// TIA Portal project "s15_motor" (V21)

(* hardware
DEVICE "S7-1500/ET200MP station_1"  S7-1500 station
   slot 0: "Rail_0"  Rack  6ES7 590-1***0-0AA0
   slot 1: "MOTORPLC"  CPU 1511-1 PN  6ES7 511-1AL03-0AB0  V4.1
      slot 3: "CPU display_1"  6ES7591-1AA00-0AA0
      slot 32768: "PROFINET interface_1"  X1
         slot 32769: "Port_1"  X1 P1
         slot 32770: "Port_2"  X1 P2
      slot 34817: "Virtual CP interface port_1"  Virtual CP interface port  Virtual CP interface port FW V4.1
*)

// ===== PLC "MOTORPLC"  CPU 1511-1 PN =====

VAR_GLOBAL   // PLC tag table "Default tag table"
   "StartPB" AT %I0.0 : Bool;   // start button, normally open
   "StopPB" AT %I0.1 : Bool;   // stop button, normally closed
   "Guard" AT %I0.2 : Bool;   // guard closed
   "MotorLadOut" AT %Q0.0 : Bool;
   "MotorSclOut" AT %Q0.1 : Bool;
END_VAR

DATA_BLOCK "MotorData"   // DB1
{ S7_Optimized_Access := 'TRUE' }
VERSION : 0.1
   VAR
      starts : Int;
      runTime : Time;
   END_VAR
BEGIN
END_DATA_BLOCK

DATA_BLOCK "MotorLAD_DB"   // DB2
{ S7_Optimized_Access := 'TRUE' }
VERSION : 0.1
// stored: InstanceOfName MotorLAD
"MotorLAD"
BEGIN
END_DATA_BLOCK

DATA_BLOCK "MotorSCL_DB"   // DB3
{ S7_Optimized_Access := 'TRUE' }
VERSION : 0.1
// stored: InstanceOfName MotorSCL
"MotorSCL"
BEGIN
END_DATA_BLOCK

FUNCTION_BLOCK "MotorLAD"   // FB1, LAD
{ S7_Optimized_Access := 'TRUE' }
VERSION : 0.1
   VAR_INPUT
      start : Bool;
      stop : Bool;
      interlock : Bool;
   END_VAR
   VAR_OUTPUT
      motor : Bool;
   END_VAR
   VAR
      run : Bool;
      runEdge : Bool;
      delay : TON_TIME;
   END_VAR
   VAR_TEMP   // added for the SCL form of the ladder/FBD networks
      _w1 : Bool;
   END_VAR
BEGIN

REGION Network 1
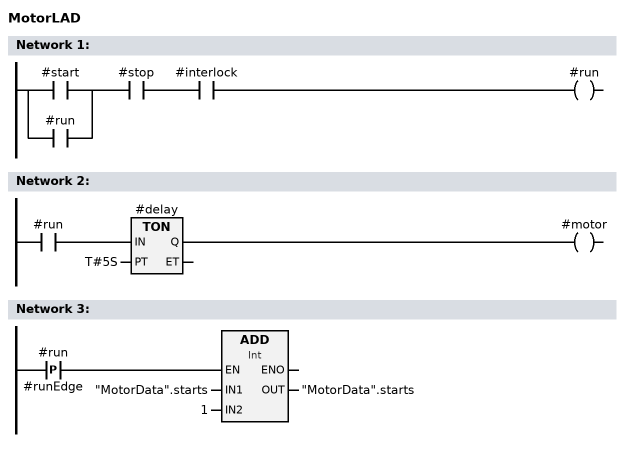
   RUNG wire#powerrail
      Contact( #start )
      wire#w1
      Contact( #stop )
      Contact( #interlock )
      Coil( #run )
   END_RUNG
   RUNG wire#powerrail
      Contact( #run )
   END_RUNG wire#w1
   // the same network as SCL:
   #run := (#start OR #run) AND #stop AND #interlock;
END_REGION

REGION Network 2
   #delay(IN := #run, PT := T#5S);   // TON
   #motor := #delay.Q;
END_REGION

REGION Network 3
   RUNG wire#powerrail
      P_Contact(operand := #run, bit := #runEdge)
      { S7_Templates := "SrcType := Int" } Add(in1 := "MotorData".starts, in2 := 1, out => "MotorData".starts)
   END_RUNG
   // the same network as SCL:
   #_w1 := #run AND NOT #runEdge;   // rising edge of #run
   #runEdge := #run;
   IF #_w1 THEN "MotorData".starts := "MotorData".starts + 1; END_IF;
END_REGION
END_FUNCTION_BLOCK

FUNCTION_BLOCK "MotorSCL"   // FB2, SCL
{ S7_Optimized_Access := 'TRUE' }
VERSION : 0.1
   VAR_INPUT
      start : Bool;
      stop : Bool;
      interlock : Bool;
   END_VAR
   VAR_OUTPUT
      motor : Bool;
   END_VAR
   VAR
      run : Bool;
      runOld : Bool;
      delay : TON_TIME;
   END_VAR
BEGIN
       // seal-in with interlock
       #run := (#start OR #run) AND #stop AND #interlock;
       // start delay
       #delay(IN := #run,
              PT := T#5S);
       #motor := #delay.Q;
       // count the starts
       IF #run AND NOT #runOld THEN
           "MotorData".starts := "MotorData".starts + 1;
       END_IF;
       #runOld := #run;
END_FUNCTION_BLOCK

ORGANIZATION_BLOCK "Main"   // OB1, LAD, ProgramCycle
TITLE = "Main Program Sweep (Cycle)"
{ S7_Optimized_Access := 'TRUE' }
VERSION : 0.1
   VAR_INPUT
      Initial_Call : Bool;   // Initial call of this OB
      Remanence : Bool;   // =True, if remanent data are available
   END_VAR
BEGIN

REGION Network 1
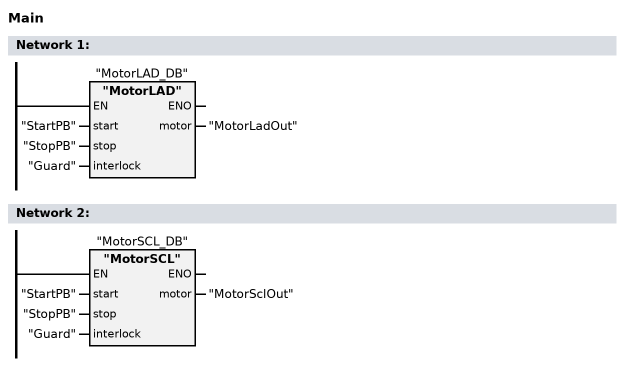
   RUNG wire#powerrail
      "MotorLAD_DB"(start := "StartPB", stop := "StopPB", interlock := "Guard", motor => "MotorLadOut")
   END_RUNG
   // the same network as SCL:
   "MotorLAD_DB"(start := "StartPB", stop := "StopPB", interlock := "Guard", motor => "MotorLadOut");   // "MotorLAD"
END_REGION

REGION Network 2
   RUNG wire#powerrail
      "MotorSCL_DB"(start := "StartPB", stop := "StopPB", interlock := "Guard", motor => "MotorSclOut")
   END_RUNG
   // the same network as SCL:
   "MotorSCL_DB"(start := "StartPB", stop := "StopPB", interlock := "Guard", motor => "MotorSclOut");   // "MotorSCL"
END_REGION
END_ORGANIZATION_BLOCK